Fanuc KAREL source: kt00018.KL

-- PROVISIONAL review KL for V1013-1; original PC SHA256 86750b30a9c7c037942d1bd22a93afb89b1c58def0900d9fc5bccdf25d838f38
-- Incomplete behavior may be omitted. Consult companion uncertainty JSON. Do not deploy.
PROGRAM KT00018
%NOLOCKGROUP
VAR
  I2 : INTEGER
  OUT : REAL
-- UNRESOLVED_DECL Y1 type=002018
BEGIN
  -- UNRESOLVED_PC offsets 5-19; opcodes 2E,22,9D,33,B2
  -- UNRESOLVED_PC offsets 24-35; opcodes 2E,23
  -- UNRESOLVED_PC offsets 40-63; opcodes 22,9D,33,B1,21,52,64,23
  -- UNRESOLVED_PC offsets 68-72; opcodes 7F
END KT00018
